// TIA Portal V21 export
// export: Created 2026-11-10T19:21:34.4655131Z, ExportSetting WithDefaults, DisplayName Totally Integrated Automation Portal, DisplayVersion V21 Update 3, DisplayName STEP 7 Professional, DisplayVersion V21 Update 3, DisplayName STEP 7 Safety, DisplayVersion V21, DisplayName Tech WebApplication, DisplayVersion V21, DisplayName WinCC Basic/Comfort/Advanced, DisplayVersion V21 Update 3, DisplayName WinCC Unified, DisplayVersion V21 Update 3
FUNCTION_BLOCK "FB_Lad_us006"   // FB10, LAD
{ S7_Optimized_Access := 'TRUE' }
VERSION : 0.1
// stored: AutoNumber true, IsIECCheckEnabled false, IsRetainMemResEnabled false, MemoryReserve 100, SetENOAutomatically false, UDAEnableTagReadback false
   VAR_INPUT
      v_req : Bool;
      v_drive : USInt;
      v_param : UInt;
      v_index : UInt;
      v_eeprom : Bool;
      v_value : P2P_USS_BASE;
   END_VAR
   VAR_OUTPUT
      v_done : Bool;
      v_error : Bool;
      v_status : Word;
   END_VAR
   VAR_IN_OUT
      v_uss_db : P2P_USS_BASE;
   END_VAR
BEGIN

REGION Network 1: USS_WPM - Change parameters in the drive
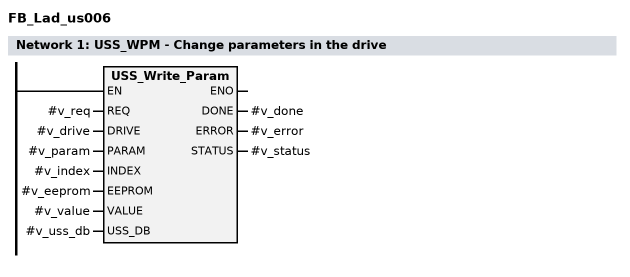
   RUNG wire#powerrail
      USS_Write_Param(REQ := #v_req, DRIVE := #v_drive, PARAM := #v_param, INDEX := #v_index, EEPROM := #v_eeprom, VALUE := #v_value, USS_DB := #v_uss_db, DONE => #v_done, ERROR => #v_error, STATUS => #v_status)
   END_RUNG
   // the same network as SCL:
   USS_Write_Param(REQ := #v_req,
                   DRIVE := #v_drive,
                   PARAM := #v_param,
                   INDEX := #v_index,
                   EEPROM := #v_eeprom,
                   VALUE := #v_value,
                   USS_DB := #v_uss_db,
                   DONE => #v_done,
                   ERROR => #v_error,
                   STATUS => #v_status);
END_REGION
END_FUNCTION_BLOCK
